// TIA Portal V20 export
Screen "200FX1Layout_Docking"  1276x673
  ScreenItem "Line_Header_X0_Y64" at 0,64 size 1276x0  Type=HmiLine
  ScreenItem "permanentareaborderrectangle" at 0,0 size 0x0  Type=HmiRectangle
  ScreenItem "Button_Back" at 2,2 size 90x60  Type=HmiButton
  ScreenItem "Move_Legend" at 1183,2 size 90x60  Type=HmiButton
  ScreenItem "Fusszeile_Button_ManualOPMode1_2" at 188,2 size 90x60  Type=HmiButton
  ScreenItem "文本域_22" at 1130,495 size 104x23  Type=HmiTextBox
  ScreenItem "面板容器_23" at 1177,528 size 96x32  Type=HmiFaceplateContainer
  ScreenItem "面板容器_22" at 1067,528 size 96x32  Type=HmiFaceplateContainer
  ScreenItem "Fusszeile_Button_ManualOPMode1_1" at 95,2 size 90x60  Type=HmiButton
  ScreenItem "LSicar_Valve8Pos_LeftHomeRightWork_WithPB_3" at 1099,110 size 160x53  Type=HmiFaceplateContainer
  ScreenItem "文本域_5" at 1107,83 size 139x22  Type=HmiTextBox
  ScreenItem "文本域_8" at 1172,-248 size 100x20  Type=HmiTextBox
  ScreenItem "文本域_9" at 1741,-563 size 100x20  Type=HmiTextBox
  ScreenItem "文本域_10" at 2310,-878 size 100x20  Type=HmiTextBox
  ScreenItem "文本域_12" at 321,1215 size 100x20  Type=HmiTextBox
  ScreenItem "Title_ScreenOverview_X390_Y2_1" at 384,2 size 510x57  Type=HmiTextBox
  ScreenItem "Button_Back_1" at 1180,606 size 90x60  Type=HmiButton
  ScreenItem "文本域_1" at -1,82 size 120x40  Type=HmiTextBox
  ScreenItem "文本域_27" at -1,126 size 120x40  Type=HmiTextBox
  ScreenItem "面板容器_2" at 1092,3 size 88x58  Type=HmiFaceplateContainer
  ScreenItem "OPMode1_Blocked" at 1166,5 size 14x14  Type=HmiGraphicView
  ScreenItem "OPMode4_Foreground_Blocked_1" at 1092,3 size 88x58  Type=HmiGraphicView
  ScreenItem "Graphic view_1" at 114,71 size 766x527  Type=HmiGraphicView
  ScreenItem "面板容器_15" at 212,527 size 65x43  Type=HmiFaceplateContainer
  ScreenItem "Line_4" at 754,235 size 166x11  Type=HmiLine
  ScreenItem "Line_5" at 784,328 size 125x31  Type=HmiLine
  ScreenItem "Line_6" at 272,381 size 237x17  Type=HmiLine
  ScreenItem "Line_7" at 292,468 size 234x64  Type=HmiLine
  ScreenItem "面板容器_13" at 913,256 size 142x51  Type=HmiFaceplateContainer
  ScreenItem "面板容器_12" at 171,410 size 142x51  Type=HmiFaceplateContainer
  ScreenItem "Faceplate container_5" at 937,365 size 65x43  Type=HmiFaceplateContainer
  ScreenItem "文本域_19" at 192,508 size 100x20  Type=HmiTextBox
  ScreenItem "文本域_6" at 172,368 size 140x40  Type=HmiTextBox
  ScreenItem "文本域_11" at 916,343 size 100x20  Type=HmiTextBox
  ScreenItem "文本域_14" at 914,214 size 140x40  Type=HmiTextBox
